Fanuc KAREL source: ko00058.KL

-- PROVISIONAL review KL for V770-1; original PC SHA256 4df20d560c78dc30e5b1ed0cff78874968f7e51f390f55db4e4f2fd55518234c
-- Incomplete behavior may be omitted. Consult companion uncertainty JSON. Do not deploy.
PROGRAM KO00058
%NOLOCKGROUP
BEGIN
  -- UNRESOLVED_PC offsets 5-12; opcodes 9D,23
  -- UNRESOLVED_PC offsets 17-69; opcodes 27,27,49,7E,AD,27,49,7E,AD,22,31,7E,4A
  -- UNRESOLVED_PC offsets 74-78; opcodes 7F
END KO00058
